// TIA Portal V21 export
// export: Created 2026-10-14T03:06:08.5383805Z, ExportSetting WithDefaults, DisplayName Totally Integrated Automation Portal, DisplayVersion V21, DisplayName STEP 7 Professional, DisplayVersion V21, DisplayName STEP 7 Safety, DisplayVersion V21, DisplayName Tech WebApplication, DisplayVersion V21, DisplayName WinCC Basic/Comfort/Advanced, DisplayVersion V21, DisplayName WinCC Unified, DisplayVersion V21
VAR_GLOBAL   // PLC tag table "Default tag table"
   SynchronousAxis_red_Actor_Interface_AddressIn AT %I260.0 : "PD_TEL105_IN";
   SynchronousAxis_red_Actor_Interface_AddressOut AT %Q260.0 : "PD_TEL105_OUT";
   PositioningAxis_blue_Actor_Interface_AddressIn AT %I280.0 : "PD_TEL105_IN";
   PositioningAxis_blue_Actor_Interface_AddressOut AT %Q280.0 : "PD_TEL105_OUT";
   Clock_Byte AT %MB0 : Byte;
   Clock_10Hz AT %M0.0 : Bool;
   Clock_5Hz AT %M0.1 : Bool;
   "Clock_2.5Hz" AT %M0.2 : Bool;
   Clock_2Hz AT %M0.3 : Bool;
   "Clock_1.25Hz" AT %M0.4 : Bool;
   Clock_1Hz AT %M0.5 : Bool;
   "Clock_0.625Hz" AT %M0.6 : Bool;
   "Clock_0.5Hz" AT %M0.7 : Bool;
END_VAR
